SUBAPPLICATION VarInOutSubappNetwork
  (* Standard: 61499-1; Description: Copyright (c) 2026 Martin Erich Jobst This program and the accompanying materials are made available under the terms of the Eclipse Public License 2.0 which is available at https://www.eclipse.org/legal/epl-2.0/ SPDX-License-Identifier: EPL-2.0 *)
  (* Version 1.0, 2026-11-18, Martin Jobst *)
  PACKAGE lib::VarDeclaration;
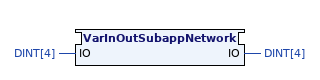
  VAR_IN_OUT
    IO : ARRAY [0..3] OF DINT;
  END_VAR
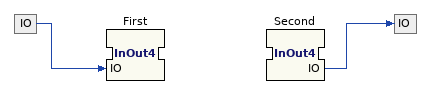
  FBS
    First : lib::VarDeclaration::support::InOut4;
    Second : lib::VarDeclaration::support::InOut4;
  END_FBS
  DATA_CONNECTIONS
    IO TO First.IO;
    Second.IO TO IO;
  END_CONNECTIONS
END_SUBAPPLICATION
